Fanuc KAREL source: KA00007.KL

PROGRAM KA00007
%NOLOCKGROUP
VAR
  SRC: INTEGER
  DST: XYZWPREXT
BEGIN
  SRC = 2
  DST = SRC
END KA00007
